DATA_BLOCK "PipDb"
{ S7_Optimized_Access := 'TRUE' }
VERSION : 0.1
NON_RETAIN
   VAR
      Ob1Count : DInt;
      Ob30Count : DInt;
   END_VAR

BEGIN

END_DATA_BLOCK

